VAR_GLOBAL
    aIn  AT %I* : ARRAY[0..15] OF BYTE;  // TxPDO 16 byte
    aOut AT %Q* : ARRAY[0..3]  OF BYTE;  // RxPDO 4 byte
END_VAR

(* stored: Version 1.1.0.1, ProductVersion 3.1.4024.16
   GVL GVL: Id {bdb62bb0-8c97-4a62-9045-c1544f9d2e00} *)
